Fanuc KAREL source: ko00066.KL

-- PROVISIONAL review KL for V1013-1; original PC SHA256 4607222923bdf6b7a1eaef20673d273b5236d5eb81cd7c8f52aa8914b391c324
-- Incomplete behavior may be omitted. Consult companion uncertainty JSON. Do not deploy.
PROGRAM KO00066
%NOLOCKGROUP
BEGIN
  -- UNRESOLVED_PC offsets 5-12; opcodes 9D,23
  -- UNRESOLVED_PC offsets 17-63; opcodes 27,22,1C,22,1C,22,31,7E,4A
  -- UNRESOLVED_PC offsets 68-72; opcodes 7F
END KO00066
